SUBAPPLICATION AuxIXA_TO_logiBUS_QXA_BG (* AUX-Funktion (Aux_IXA) auf DigitalOutput QXA mit GreenWhiteBackground. Generisch, analog zu Button_IXA_TO_logiBUS_QXA_BG (dort Button statt AUX). *)
  (* Standard: 61499-2 *)
  (* Version 1.0, 2026-09-09, Franz Höpfinger, Meisterschulen am Ostbahnhof, Ausgelagert aus Uebung_010f2_sub_AX zur Wiederverwendung. *)
  PACKAGE MyLib::sys;
  IMPORT isobus::UT::Q::const::IDs::ID_NULL;
  IMPORT logiBUS::io::DQ::logiBUS_DO;
  IMPORT logiBUS::io::DQ::logiBUS_DO_S;
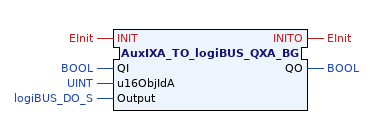
  EVENT_INPUT
    INIT : EInit; (* Initialization Request *)
  END_EVENT
  EVENT_OUTPUT
    INITO : EInit; (* Initialization Confirm *)
  END_EVENT
  VAR_INPUT
    QI : BOOL := TRUE; (* Quality Input - TRUE to enable service *)
    u16ObjIdA : UINT := ID_NULL; (* Object ID AUX *)
    Output : logiBUS::io::DQ::logiBUS_DO_S := logiBUS_DO::Invalid; (* Identify the Output Output_Q1..Q8 *)
  END_VAR
  VAR_OUTPUT
    QO : BOOL; (* Quality Output - TRUE if service executed successfully *)
  END_VAR
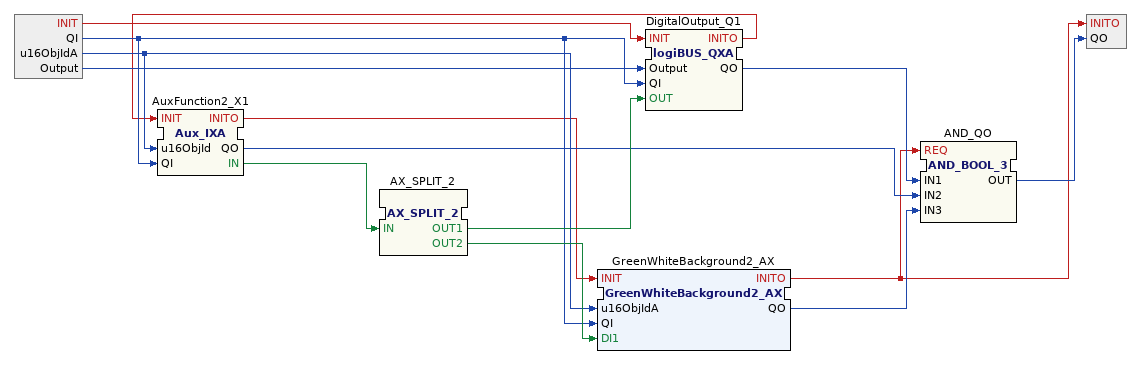
  FBS
    DigitalOutput_Q1 : logiBUS::io::DQ::logiBUS_QXA;
    AuxFunction2_X1 : isobus::UT::io::Auxiliary::IN::Aux_IXA;
    AX_SPLIT_2 : adapter::events::unidirectional::AX_SPLIT_2;
    AND_QO : iec61131::booleanOperators::AND_BOOL_3;
  END_FBS
  SUBAPPS
    GreenWhiteBackground2_AX : MyLib::sys::GreenWhiteBackground2_AX;
  END_SUBAPPS
  EVENT_CONNECTIONS
    INIT TO DigitalOutput_Q1.INIT;
    DigitalOutput_Q1.INITO TO AuxFunction2_X1.INIT;
    AuxFunction2_X1.INITO TO GreenWhiteBackground2_AX.INIT;
    GreenWhiteBackground2_AX.INITO TO INITO;
    GreenWhiteBackground2_AX.INITO TO AND_QO.REQ;
  END_CONNECTIONS
  DATA_CONNECTIONS
    u16ObjIdA TO AuxFunction2_X1.u16ObjId;
    u16ObjIdA TO GreenWhiteBackground2_AX.u16ObjIdA;
    Output TO DigitalOutput_Q1.Output;
    QI TO DigitalOutput_Q1.QI;
    QI TO AuxFunction2_X1.QI;
    DigitalOutput_Q1.QO TO AND_QO.IN1;
    AuxFunction2_X1.QO TO AND_QO.IN2;
    AND_QO.OUT TO QO;
    QI TO GreenWhiteBackground2_AX.QI;
    GreenWhiteBackground2_AX.QO TO AND_QO.IN3;
  END_CONNECTIONS
  ADAPTER_CONNECTIONS
    AuxFunction2_X1.IN TO AX_SPLIT_2.IN;
    AX_SPLIT_2.OUT1 TO DigitalOutput_Q1.OUT;
    AX_SPLIT_2.OUT2 TO GreenWhiteBackground2_AX.DI1;
  END_CONNECTIONS
END_SUBAPPLICATION
